(* IEC 61131-3 sources: volt/packages/volt-lsp-iec/test-corpus/pro2193/Device/Plc Logic/Application/01 Main/IQ Handling/Data, 5 files *)

(* ---- Slice_Type.dut ---- *)
TYPE Slice_Type :
STRUCT
	sliceName	: STRING(40);
	isOutput	: BOOL;
	component	: ARRAY[1..8] OF SliceComponent_Type;
END_STRUCT
END_TYPE

(* ---- SliceComponent_Type.dut ---- *)
TYPE SliceComponent_Type :
STRUCT
	name		: STRING(80);
	actValue	: BOOL;
	forceValue	: BOOL;
END_STRUCT
END_TYPE

(* ---- MapperBase.pou ---- *)
FUNCTION_BLOCK INTERNAL ABSTRACT MapperBase
VAR_INPUT
	sliceNumber		: IQSlices;
END_VAR
VAR
	sliceInfo		: REFERENCE TO Slice_Type;
	sliceForced		: REFERENCE TO BOOL;
	i				: INT;
END_VAR

%LANGUAGE ST
IF __ISVALIDREF(sliceInfo) THEN
	sliceInfo.sliceName		:= TO_STRING(sliceNumber);
END_IF

END_FUNCTION_BLOCK

METHOD PUBLIC SetSliceRef
VAR_INPUT
	sliceInfo	: REFERENCE TO Slice_Type;
	sliceForced	: REFERENCE TO BOOL;
END_VAR

%LANGUAGE ST
THIS^.sliceInfo		REF= sliceInfo;
THIS^.sliceForced	REF= sliceForced;

END_METHOD

(* ---- MapperInputs.pou ---- *)
// Mapping digital inputs. Use to map a byte into 8 individual bits
FUNCTION_BLOCK INTERNAL MapperInputs
EXTENDS MapperBase
VAR_INPUT
	slice			: REFERENCE TO BYTE;
END_VAR
VAR_OUTPUT
	bit1			: BIT;
	bit2			: BIT;
	bit3			: BIT;
	bit4			: BIT;
	bit5			: BIT;
	bit6			: BIT;
	bit7			: BIT;
	bit8			: BIT;
END_VAR

%LANGUAGE ST
SUPER^();

IF __ISVALIDREF(sliceInfo) THEN
	sliceInfo.isOutput					:= FALSE;
	FOR i := 1 TO 8 DO
		sliceInfo.component[i].name		:= GVL_IQ.inputs[sliceNumber][i];
		sliceInfo.component[i].actValue	:= BitLogic.ExtractFromByte(slice, TO_BYTE(i-1));
	END_FOR
END_IF

bit1	:= slice.0;
bit2	:= slice.1;
bit3	:= slice.2;
bit4	:= slice.3;
bit5	:= slice.4;
bit6	:= slice.5;
bit7	:= slice.6;
bit8	:= slice.7;

END_FUNCTION_BLOCK

(* ---- MapperOutputs.pou ---- *)
// Mapping digital outputs. Use to map 8 individual bits into a byte
FUNCTION_BLOCK INTERNAL MapperOutputs
EXTENDS MapperBase
VAR_INPUT
	slice			: REFERENCE TO BYTE;
	bit1			: BIT;
	bit2			: BIT;
	bit3			: BIT;
	bit4			: BIT;
	bit5			: BIT;
	bit6			: BIT;
	bit7			: BIT;
	bit8			: BIT;
END_VAR

%LANGUAGE ST
SUPER^();

IF __ISVALIDREF(sliceForced) AND_THEN sliceForced THEN
	slice.0	:= sliceInfo.component[1].forceValue;
	slice.1	:= sliceInfo.component[2].forceValue;
	slice.2	:= sliceInfo.component[3].forceValue;
	slice.3	:= sliceInfo.component[4].forceValue;
	slice.4	:= sliceInfo.component[5].forceValue;
	slice.5	:= sliceInfo.component[6].forceValue;
	slice.6	:= sliceInfo.component[7].forceValue;
	slice.7	:= sliceInfo.component[8].forceValue;
ELSE
	slice.0	:= bit1;
	slice.1	:= bit2;
	slice.2	:= bit3;
	slice.3	:= bit4;
	slice.4	:= bit5;
	slice.5	:= bit6;
	slice.6	:= bit7;
	slice.7	:= bit8;
END_IF

IF __ISVALIDREF(sliceInfo) THEN
	sliceInfo.isOutput					:= TRUE;
	FOR i := 1 TO 8 DO
		sliceInfo.component[i].name		:= GVL_IQ.outputs[sliceNumber][i];
		sliceInfo.component[i].actValue	:= BitLogic.ExtractFromByte(slice, TO_BYTE(i-1));
	END_FOR
END_IF

END_FUNCTION_BLOCK
